(* IEC 61131-3 sources: Twinova/app/src-tauri/project/tests/fixtures/invalid/duplicate_id/components, 3 files *)

(* ---- twinova.belt@1.st ---- *)
(* Twinova belt conveyor, its drive, re-expressed from Open Industry Project's conveyor drive
   (examples/parts/_shared/conveyorDrive.js at 1e7488c, MIT). While the PLC's run is on, the surface ramps to
   speed_ref, which reads the speed parameter unless the PLC writes it: up at speed_at_30 per accel_time, down at
   speed_at_30 per decel_time, through 0 before it reverses; a ramp time of 0 is instant. running reports run after
   the start delay. The conveyor's native model reads surface_speed, and publishes the velocity, the encoder and the
   pulse itself. The field cycles every 1 ms, and TIME_TO_DWORD gives whole milliseconds, made a REAL through DINT:
   truST's DWORD_TO_REAL keeps the bits, not the number. n steps of speed_at_30 / n add up to speed_at_30 only within
   a rounding of REAL, so the ramp lands on its target within a hundredth of a step, on its millisecond. At its
   target the ramp is skipped. *)
FUNCTION_BLOCK BeltBehaviour
VAR_INPUT
    start_delay : TIME;
    accel_time : TIME;
    decel_time : TIME;
    speed_at_30 : REAL;
END_VAR
VAR_OUTPUT
    surface_speed : REAL;
END_VAR
VAR
    run AT %I* : BOOL;
    speed_ref AT %I* : REAL;
    running AT %Q* : BOOL;
    started : TON;
    target : REAL;
    ramp : TIME;
    step : REAL;
END_VAR
IF run THEN
    target := speed_ref;
ELSE
    target := 0.0;
END_IF;
IF target <> surface_speed THEN
    IF target * surface_speed < 0.0 THEN
        IF decel_time > T#0MS THEN
            target := 0.0;
        ELSE
            surface_speed := 0.0;
        END_IF;
    END_IF;
    IF ABS(target) > ABS(surface_speed) THEN
        ramp := accel_time;
    ELSE
        ramp := decel_time;
    END_IF;
    step := 0.0;
    IF ramp > T#0MS THEN
        step := speed_at_30 / DINT_TO_REAL(DWORD_TO_DINT(TIME_TO_DWORD(ramp)));
    END_IF;
    IF step <= 0.0 OR ABS(target - surface_speed) <= step * 1.01 THEN
        surface_speed := target;
    ELSIF target > surface_speed THEN
        surface_speed := surface_speed + step;
    ELSE
        surface_speed := surface_speed - step;
    END_IF;
END_IF;
started(IN := run, PT := start_delay);
running := started.Q;
END_FUNCTION_BLOCK

(* ---- twinova.chain_transfer@1.st ---- *)
(* Twinova chain transfer, re-expressed from Open Industry Project's chain transfer
   (examples/parts/chain-transfer/behavior.ts at 1e7488c, MIT). popup raises the chains and carries sideways at once;
   the lift slews linearly over raise_time, as OIP's approach(). raised_fb reports the top of the stroke, which OIP
   does not have. The field cycles every 1 ms (spec 2026-11-09-component-behaviour-design.md, decision 3), so travel
   counts the milliseconds of stroke done; TIME_TO_DWORD gives whole milliseconds. *)
FUNCTION_BLOCK ChainTransferBehaviour
VAR_INPUT
    raise_time : TIME;
END_VAR
VAR_OUTPUT
    lift : REAL;
    raised : BOOL;
END_VAR
VAR
    popup AT %I* : BOOL;
    raised_fb AT %Q* : BOOL;
    stroke : DINT;
    travel : DINT;
END_VAR
raised := popup;
stroke := MAX(DWORD_TO_DINT(TIME_TO_DWORD(raise_time)), 1);
IF raised THEN
    travel := MIN(travel + 1, stroke);
ELSE
    travel := MAX(travel - 1, 0);
END_IF;
lift := DINT_TO_REAL(travel) / DINT_TO_REAL(stroke);
raised_fb := raised AND travel = stroke;
END_FUNCTION_BLOCK

(* ---- twinova.roller@1.st ---- *)
(* Twinova roller conveyor, its drive, re-expressed from Open Industry Project's conveyor drive
   (examples/parts/_shared/conveyorDrive.js at 1e7488c, MIT). While the PLC's run is on, the surface ramps to
   speed_ref, which reads the speed parameter unless the PLC writes it: up at speed_at_30 per accel_time, down at
   speed_at_30 per decel_time, through 0 before it reverses; a ramp time of 0 is instant. running reports run after
   the start delay. The conveyor's native model reads surface_speed, and publishes the velocity, the encoder and the
   pulse itself. The field cycles every 1 ms, and TIME_TO_DWORD gives whole milliseconds, made a REAL through DINT:
   truST's DWORD_TO_REAL keeps the bits, not the number. n steps of speed_at_30 / n add up to speed_at_30 only within
   a rounding of REAL, so the ramp lands on its target within a hundredth of a step, on its millisecond. At its
   target the ramp is skipped. *)
FUNCTION_BLOCK RollerBehaviour
VAR_INPUT
    start_delay : TIME;
    accel_time : TIME;
    decel_time : TIME;
    speed_at_30 : REAL;
END_VAR
VAR_OUTPUT
    surface_speed : REAL;
END_VAR
VAR
    run AT %I* : BOOL;
    speed_ref AT %I* : REAL;
    running AT %Q* : BOOL;
    started : TON;
    target : REAL;
    ramp : TIME;
    step : REAL;
END_VAR
IF run THEN
    target := speed_ref;
ELSE
    target := 0.0;
END_IF;
IF target <> surface_speed THEN
    IF target * surface_speed < 0.0 THEN
        IF decel_time > T#0MS THEN
            target := 0.0;
        ELSE
            surface_speed := 0.0;
        END_IF;
    END_IF;
    IF ABS(target) > ABS(surface_speed) THEN
        ramp := accel_time;
    ELSE
        ramp := decel_time;
    END_IF;
    step := 0.0;
    IF ramp > T#0MS THEN
        step := speed_at_30 / DINT_TO_REAL(DWORD_TO_DINT(TIME_TO_DWORD(ramp)));
    END_IF;
    IF step <= 0.0 OR ABS(target - surface_speed) <= step * 1.01 THEN
        surface_speed := target;
    ELSIF target > surface_speed THEN
        surface_speed := surface_speed + step;
    ELSE
        surface_speed := surface_speed - step;
    END_IF;
END_IF;
started(IN := run, PT := start_delay);
running := started.Q;
END_FUNCTION_BLOCK
